// TIA Portal V21 export
// export: Created 2026-11-07T15:50:59.7595138Z, ExportSetting WithDefaults, DisplayName Totally Integrated Automation Portal, DisplayVersion V21, DisplayName STEP 7 Professional, DisplayVersion V21, DisplayName STEP 7 Safety, DisplayVersion V21, DisplayName Tech WebApplication, DisplayVersion V21, DisplayName WinCC Basic/Comfort/Advanced, DisplayVersion V21, DisplayName WinCC Unified, DisplayVersion V21
TextList "TL_Bay"  ListRange=Decimal
  TextListEntry   EntryType=SingleValue, Text="0 BROD"
  TextListEntry   EntryType=SingleValue, From=1, To=1, Text="1 SKLADIŠTE"
